KUKA KRL data list: folge125.dat

&ACCESS RVP
&REL 1
&COMMENT bt2krl sim data Folge 125 plan 16#A312
DEFDAT FOLGE125
   ; Generated by bt2krl 0.1.0 from bt2plc plan bt_1791274820_cell_2robot (cell cell_2robot), PLAN_ID 16#A312
   ; Robot robot1 (R1), controller robot1, model KR240R2900_ULTRA, joint mapping identity
   ; Profile sim (bt2plc simulator telegram). NEVER install on a VW KS24 robot:
   ; its signals collide with the VW standard (Fertigmeldung, interlocks, PRG_NR).
   ; Do not edit: regenerate with bt2krl (plain KRL, no inline forms).
   EXT BAS (BAS_COMMAND :IN,REAL :IN )
   DECL AXIS PHOME={A1 0.0,A2 -90.0,A3 90.0,A4 0.0,A5 0.0,A6 0.0}
ENDDAT
